// TIA Portal V21 export
// export: Created 2026-11-10T07:35:08.5503435Z, ExportSetting WithDefaults, DisplayName Totally Integrated Automation Portal, DisplayVersion V21 Update 3, DisplayName STEP 7 Professional, DisplayVersion V21 Update 3, DisplayName STEP 7 Safety, DisplayVersion V21, DisplayName Tech WebApplication, DisplayVersion V21, DisplayName WinCC Basic/Comfort/Advanced, DisplayVersion V21 Update 3, DisplayName WinCC Unified, DisplayVersion V21 Update 3
FUNCTION_BLOCK "FB_Lad_ex065"   // FB68, LAD
{ S7_Optimized_Access := 'TRUE' }
VERSION : 0.1
// stored: AutoNumber true, IsIECCheckEnabled false, IsRetainMemResEnabled false, MemoryReserve 100, SetENOAutomatically false, UDAEnableTagReadback false
   VAR_INPUT
      v_req : Bool;
      v_laddr : HW_DPSLAVE;
      v_ret_val : DInt;
   END_VAR
   VAR_OUTPUT
      v_busy : Bool;
   END_VAR
   VAR_IN_OUT
      v_record : Variant;
   END_VAR
BEGIN

REGION Network 1: DPNRM_DG - Read diagnostics data from a DP slave
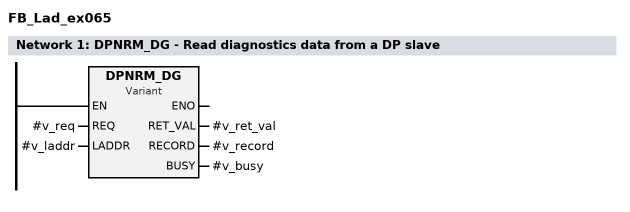
   RUNG wire#powerrail
      { S7_Templates := "[ptr_type := Variant, laddr_type := HW_DPSLAVE]" } DPNRM_DG(REQ := #v_req, LADDR := #v_laddr, RET_VAL => #v_ret_val, RECORD => #v_record, BUSY => #v_busy)
   END_RUNG
   // the same network as SCL:
   #v_ret_val := DPNRM_DG(REQ := #v_req, LADDR := #v_laddr, RECORD => #v_record, BUSY => #v_busy);
END_REGION
END_FUNCTION_BLOCK
